{attribute 'qualified_only'}
{attribute 'strict'}
TYPE
    eTcoLoggerTests :
    (
		PushMessage := 10,
		PushMessageMultiple := 20,
		PushMessageMultipleInMoreCycles := 30,
		SimplePush := 40		
    );
END_TYPE

(* stored: Version 1.1.0.1
   DUT eTcoLoggerTests: Id {3152a930-9ddc-047f-03f1-d36a10a1ade6} *)
